// Mitsubishi GX Works2 project: Task2_Ex_4   PLC: FX3G

PROGRAM MAIN
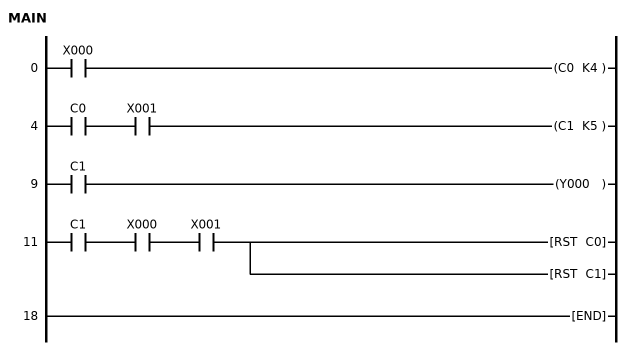
0     LD      X000
      OUT     C0 K4
4     LD      C0
      AND     X001
      OUT     C1 K5
9     LD      C1
      OUT     Y000
11    LD      C1
      AND     X000
      AND     X001
      RST     C0
      RST     C1
18    END
END_PROGRAM
